(* IEC 61131-3 sources: llm-plc-st-eval/data/processed_definitivo/gemini-3.1-pro-preview/B8/few_shot, 3 files *)

(* ---- ejec_1.st ---- *)
FUNCTION_BLOCK FB_Puerta
VAR_INPUT
    puertaAbierta : BOOL; (* Señal de puerta abierta *)
    reset : BOOL; (* Reset del registro *)
END_VAR
VAR_OUTPUT
    aviso : BOOL; (* Aviso por 5 o mas aperturas *)
    nAperturas : INT; (* Contador de aperturas *)
END_VAR
VAR
    contador : CTU; (* Contador ascendente *)
END_VAR

(* Cuenta los flancos de subida y activa el aviso al llegar a 5 *)
contador(CU := puertaAbierta, RESET := reset, PV := 5);
aviso := contador.Q;
nAperturas := contador.CV;
END_FUNCTION_BLOCK

(* ---- ejec_2.st ---- *)
FUNCTION_BLOCK FB_Puerta
VAR_INPUT
    puertaAbierta : BOOL; (* Senal de puerta abierta *)
    reset : BOOL; (* Resetea el contador y el aviso *)
END_VAR
VAR_OUTPUT
    aviso : BOOL; (* Aviso de 5 o mas aperturas *)
    nAperturas : INT; (* Numero de aperturas registradas *)
END_VAR
VAR
    flancoApertura : R_TRIG; (* Detector de flanco ascendente *)
END_VAR

(* Deteccion de transicion de FALSE a TRUE *)
flancoApertura(CLK := puertaAbierta);

(* Logica de reseteo e incremento del contador *)
IF reset THEN
    nAperturas := 0;
ELSIF flancoApertura.Q THEN
    nAperturas := nAperturas + 1;
END_IF;

(* Activacion del aviso al acumular 5 o mas aperturas *)
aviso := (nAperturas >= 5);
END_FUNCTION_BLOCK

(* ---- ejec_3.st ---- *)
FUNCTION_BLOCK FB_Puerta
VAR_INPUT
    puertaAbierta : BOOL; (* Señal de puerta abierta *)
    reset : BOOL; (* Reinicia el registro y el aviso *)
END_VAR
VAR_OUTPUT
    aviso : BOOL; (* Activo al alcanzar 5 o mas aperturas *)
    nAperturas : INT; (* Contador de aperturas *)
END_VAR
VAR
    flancoApertura : R_TRIG; (* Detector de flanco de subida *)
END_VAR

(* Deteccion de la transicion de FALSE a TRUE *)
flancoApertura(CLK := puertaAbierta);

(* Logica de reinicio y conteo *)
IF reset THEN
    nAperturas := 0;
ELSIF flancoApertura.Q THEN
    nAperturas := nAperturas + 1;
END_IF;

(* Evaluacion del aviso *)
aviso := (nAperturas >= 5);
END_FUNCTION_BLOCK
